DATA_BLOCK "FRK_SetRuntime"
{ S7_Optimized_Access := 'TRUE' }
VERSION : 0.1
NON_RETAIN
VAR
    Work {ExternalAccessible := 'False'; ExternalVisible := 'False'; ExternalWritable := 'False'} : Array[1..1] of "FRK_SetWorkspace";
END_VAR
BEGIN
END_DATA_BLOCK
